Staubli VAL3: PgProg.pjx

--- PgProg.pjx ---
Parameters version=s7.5.3 stackSize=5000 millimeterUnit=true
Program file=MoveJoint.pgx
Program file=MoveLine.pgx
Program file=MoveCirc.pgx
Program file=start.pgx
Program file=stop.pgx
Program file=main.pgx
Data file=PgProg.dtx

--- PgProg.dtx ---
mdesc mNomSpeed
frame fFrame1 = {x=1234.570, y=-98.765, z=50.500, rx=-0.000, ry=0.000, rz=30.000, fatherId=world[0]}
dio Input[16]
  [0] = {link=BasicIO-1\%I0}
  [1] = {link=BasicIO-1\%I1}
  [2] = {link=BasicIO-1\%I2}
  [3] = {link=BasicIO-1\%I3}
  [4] = {link=BasicIO-1\%I4}
  [5] = {link=BasicIO-1\%I5}
  [6] = {link=BasicIO-1\%I6}
  [7] = {link=BasicIO-1\%I7}
  [8] = {link=BasicIO-1\%I8}
  [9] = {link=BasicIO-1\%I9}
  [10] = {link=BasicIO-1\%I10}
  [11] = {link=BasicIO-1\%I11}
  [12] = {link=BasicIO-1\%I12}
  [13] = {link=BasicIO-1\%I13}
  [14] = {link=BasicIO-1\%I14}
  [15] = {link=BasicIO-1\%I15}
dio Output[16]
  [0] = {link=BasicIO-1\%Q0}
  [1] = {link=BasicIO-1\%Q1}
  [2] = {link=BasicIO-1\%Q2}
  [3] = {link=BasicIO-1\%Q3}
  [4] = {link=BasicIO-1\%Q4}
  [5] = {link=BasicIO-1\%Q5}
  [6] = {link=BasicIO-1\%Q6}
  [7] = {link=BasicIO-1\%Q7}
  [8] = {link=BasicIO-1\%Q8}
  [9] = {link=BasicIO-1\%Q9}
  [10] = {link=BasicIO-1\%Q10}
  [11] = {link=BasicIO-1\%Q11}
  [12] = {link=BasicIO-1\%Q12}
  [13] = {link=BasicIO-1\%Q13}
  [14] = {link=BasicIO-1\%Q14}
  [15] = {link=BasicIO-1\%Q15}
tool tCurrentTool = {x=0.000, y=0.000, z=200.000, rx=-0.000, ry=0.000, rz=-0.000, fatherId=flange[0], ioLink=ValveIO/valve1}
mdesc mCurrentSpeed
pointRx pPointRx = {fatherId=fFrame1[0]}
pointRx pPointRx2 = {fatherId=fFrame1[0]}

--- main.pgx ---
program main()
begin
  close(tCurrentTool)
  pPointRx.config.shoulder = lefty
  pPointRx.config.elbow = epositive
  pPointRx.config.wrist = wpositive
  pPointRx2.config.shoulder = lefty
  pPointRx2.config.elbow = epositive
  pPointRx2.config.wrist = wpositive
  mCurrentSpeed.tvel = 100.00
  mCurrentSpeed.blend = joint
  mCurrentSpeed.reach = 0.010
  mCurrentSpeed.leave = 0.010
  // Program PgProg start
  // Program generated by RoboDK v6.0.7 for Staubli RX130B on XX/XX/XXXX 18:00:00
  // Using nominal kinematics.
  mCurrentSpeed.tvel = 250.000
  mCurrentSpeed.reach = 5.000
  mCurrentSpeed.leave = 5.000
  call MoveJoint(0.00000,-10.00000,20.00000,0.00000,30.00000,0.00000)
  call MoveLine(-607.850,543.849,363.215,136.262,30.757,-130.375)
  call MoveCirc(-602.951,596.788,316.595,136.262,30.757,-130.375,-663.517,575.988,286.611,136.262,30.757,-130.375)
  call MoveJoint(20.00000,-10.00000,20.00000,0.00000,30.00000,0.00000)
  mCurrentSpeed.tvel = 100.000
  call MoveLine(-650.861,503.437,361.399,136.262,30.757,-130.375)
  mCurrentSpeed.reach = 0.000
  mCurrentSpeed.leave = 0.000
  call MoveLine(-640.584,506.980,371.534,136.262,30.757,-130.375)
  delay(0.500)
  popUpMsg("Paused. Press OK to continue")
  popUpMsg("Hello from postgen")
  // a comment
  //call prog:SubProgram()
  CustomCode(42)
  ThreadProg
  Output[1]=true
  Valve=false
  Output[3]=2.5
  watch(Input[2]==true)
  watch(Input[4]==false,1500.0)
  call MoveJoint(0.00000,-10.00000,20.00000,0.00000,30.00000,0.00000)
  call MoveJoint(10.00000,-5.00000,25.00000,5.00000,35.00000,5.00000)
  call MoveLine(-353.026,-90.135,331.702,164.619,39.324,-168.579)

  waitEndMove()
  // Program PgProg end

end

--- start.pgx ---
program start()
begin
  call main()
end

--- MoveCirc.pgx ---
program MoveCirc(num x_nX, num x_nY, num x_nZ, num x_nRx, num x_nRy, num x_nRz, num x_nX2, num x_nY2, num x_nZ2, num x_nRx2, num x_nRy2, num x_nRz2)
begin
  pPointRx.trsf.x = x_nX
  pPointRx.trsf.y = x_nY
  pPointRx.trsf.z = x_nZ
  pPointRx.trsf.rx = x_nRx
  pPointRx.trsf.ry = x_nRy
  pPointRx.trsf.rz = x_nRz
  pPointRx2.trsf.x = x_nX2
  pPointRx2.trsf.y = x_nY2
  pPointRx2.trsf.z = x_nZ2
  pPointRx2.trsf.rx = x_nRx2
  pPointRx2.trsf.ry = x_nRy2
  pPointRx2.trsf.rz = x_nRz2
  movec(pPointRx,pPointRx2,tCurrentTool,mCurrentSpeed)
end

--- MoveJoint.pgx ---
program MoveJoint(num x_nJ1, num x_nJ2, num x_nJ3, num x_nJ4, num x_nJ5, num x_nJ6)
  local joint l_jJoint
begin
  l_jJoint.j1 = x_nJ1
  l_jJoint.j2 = x_nJ2
  l_jJoint.j3 = x_nJ3
  l_jJoint.j4 = x_nJ4
  l_jJoint.j5 = x_nJ5
  l_jJoint.j6 = x_nJ6
  movej(l_jJoint,tCurrentTool ,mCurrentSpeed)
end

--- MoveLine.pgx ---
program MoveLine(num x_nX, num x_nY, num x_nZ, num x_nRx, num x_nRy, num x_nRz)
begin
  pPointRx.trsf.x = x_nX
  pPointRx.trsf.y = x_nY
  pPointRx.trsf.z = x_nZ
  pPointRx.trsf.rx = x_nRx
  pPointRx.trsf.ry = x_nRy
  pPointRx.trsf.rz = x_nRz
  movel(pPointRx,tCurrentTool,mCurrentSpeed)
end

--- stop.pgx ---
program stop()
begin
end
